(* IEC 61131-3 sources: llm-plc-st-eval/data/definitivo/gemini-3.1-pro-preview/B1/few_shot, 3 files *)

(* ---- ejec_1.st ---- *)
FUNCTION_BLOCK FB_Motor
VAR_INPUT
    btnMarcha : BOOL; (* Boton de marcha *)
    btnParo : BOOL;   (* Boton de paro *)
    btnEmerg : BOOL;  (* Paro de emergencia *)
END_VAR
VAR_OUTPUT
    motorOn : BOOL;   (* Estado del motor *)
END_VAR
VAR
    trigMarcha : R_TRIG; (* Detector de flanco para evitar rearranque *)
END_VAR

(* Detecta el flanco de subida de la marcha para que no rearranque si se mantiene pulsado *)
trigMarcha(CLK := btnMarcha);

(* Enclavamiento del motor con prioridad a las señales de paro *)
motorOn := (motorOn OR trigMarcha.Q) AND NOT btnParo AND NOT btnEmerg;
END_FUNCTION_BLOCK

(* ---- ejec_2.st ---- *)
FUNCTION_BLOCK FB_Motor
VAR_INPUT
    btnMarcha : BOOL; (* Boton de marcha *)
    btnParo : BOOL;   (* Boton de paro normal *)
    btnEmerg : BOOL;  (* Boton de paro de emergencia *)
END_VAR
VAR_OUTPUT
    motorOn : BOOL;   (* Estado de activacion del motor *)
END_VAR
VAR
    flancoMarcha : R_TRIG; (* Detector de flanco para evitar rearranque accidental *)
END_VAR

(* Detecta solo el instante en que se pulsa la marcha *)
flancoMarcha(CLK := btnMarcha);

(* Logica de enclavamiento: prioridad a las senales de paro *)
IF btnParo OR btnEmerg THEN
    motorOn := FALSE;
ELSIF flancoMarcha.Q THEN
    motorOn := TRUE;
END_IF;
END_FUNCTION_BLOCK

(* ---- ejec_3.st ---- *)
FUNCTION_BLOCK FB_Motor
VAR_INPUT
    btnMarcha : BOOL; (* Boton de marcha *)
    btnParo : BOOL;   (* Boton de paro normal *)
    btnEmerg : BOOL;  (* Boton de paro de emergencia *)
END_VAR
VAR_OUTPUT
    motorOn : BOOL;   (* Estado de activacion del motor *)
END_VAR
VAR
    flancoMarcha : R_TRIG; (* Detector de flanco para evitar rearranque *)
END_VAR

(* Detecta solo el instante en que se presiona el boton de marcha *)
flancoMarcha(CLK := btnMarcha);

(* Logica de enclavamiento con prioridad a las señales de paro *)
motorOn := (motorOn OR flancoMarcha.Q) AND NOT (btnParo OR btnEmerg);
END_FUNCTION_BLOCK
